{attribute 'qualified_only'}
//{attribute 'strict'}
{attribute 'to_string'}
TYPE E_Element_State_Long :
(
eOff := 0,
eStandby,
eNotClean,
eCIP_1_Rinzed,
eCIP_2_Deterged,
eCIP_3_Deterged_Clean,
eCIP_4_Sanitized,
eCIP_5_Done,
eWaterReady,
eReady,
eProduction,
// jump to eReady
eEmpty,
eExpired
);
END_TYPE

(* stored: Version 1.1.0.1, ProductVersion 3.1.4024.12
   DUT E_Element_State_Long: Id {d33f2c3d-ac0d-4e03-9911-2c0fb1f656b1} *)
